{attribute 'qualified_only'}
VAR_GLOBAL
    fbTempWarning  : FB_TcAlarm;
	fbPressWarning : FB_TcAlarm;
	fbTempTrip     : FB_TcAlarm;
	fbPressTrip    : FB_TcAlarm;
	fbEstop        : FB_TcAlarm;
END_VAR

(* stored: Version 1.1.0.1, ProductVersion 3.1.4026.21
   GVL gAL: Id {2cdc2925-fe36-4f2d-bd9e-9a13bda012f8} *)
